GLOBALCONSTANTS Diag (* Konstanten für Übung 141 (DiagSetDTC, Drahtbruch AI6) *)
  (* Standard: 61499-1; Description: Copyright (c) 2026 Meisterschulen am Ostbahnhof This program and the accompanying materials are made available under the terms of the Eclipse Public License 2.0 which is available at https://www.eclipse.org/legal/epl-2.0/ SPDX-License-Identifier: EPL-2.0 *)
  (* Version 1.0, 2026-11-17, Franz Höpfinger, Meisterschulen am Ostbahnhof, Drahtbruch 4-20 mA als DTC *)
  PACKAGE Uebungen::const::Uebung_140_149;
  VAR_GLOBAL CONSTANT
    SPN_DRAHTBRUCH_AI6 : UDINT := 520192; (* 141: erster proprietärer SPN (J1939DA) *)
    MV_DRAHTBRUCH : UDINT := 564; (* 141: unter 564 mV (3,6 mA) = Drahtbruch *)
    MV_OK : UDINT := 626; (* 141: ab 626 mV (4 mA) wieder OK *)
  END_VAR
END_GLOBALCONSTANTS
